(* IEC 61131-3 sources: kns-port-domestic/targets/astra/src/POUs/Model/F_PumpCurrent, 2 files *)

(* ---- F_PumpCurrent.decl.st ---- *)
// Назначение: ток двигателя насоса в модели, А. Гидравлическая мощность
//             P_hyd = ρ·g·(q/3600)·H/1000 кВт; потребляемая P = max(P_hyd/η, rLossShare·Pnom·s³) —
//             не меньше потерь без подачи, поэтому ток непрерывен при закрытии обратного клапана;
//             I = rImagShare·Inom·s + (1 − rImagShare)·Inom·P/Pnom. Без вращения (s ≤ 0), при
//             неверной характеристике или неконечных входах — 0.
// Автор:      kr0nsch
// Версия:     0.1.0
// Документ:   docs/DESIGN.md, разделы 11.2, 11.3
FUNCTION F_PumpCurrent : REAL
VAR_INPUT
    rFlow_m3h : REAL;           // подача насоса
    rHead_m   : REAL;           // напор сети в рабочей точке
    rSpeed    : REAL;           // относительная скорость s = f / 50 Гц
    stPump    : ST_PumpModelCfg;  // характеристика насоса и двигателя
END_VAR
VAR
    rHyd_kW  : REAL;            // гидравлическая мощность
    rLoss_kW : REAL;            // потери без подачи
    rIn_kW   : REAL;            // потребляемая мощность
END_VAR

(* ---- F_PumpCurrent.impl.st ---- *)
F_PumpCurrent := 0.0;
IF NOT (PL.F_IsFinite(rIn := rFlow_m3h) AND PL.F_IsFinite(rIn := rHead_m) AND PL.F_IsFinite(rIn := rSpeed)) THEN
    RETURN;
END_IF
IF rSpeed <= 0.0 OR stPump.rPnom_kW <= 0.0 OR stPump.rEta <= 0.0 THEN
    RETURN;
END_IF

rHyd_kW := GVL_Const.SIM_RHO_KGM3 * GVL_Const.SIM_GRAVITY_MPS2 * (MAX(rFlow_m3h, 0.0) / GVL_Const.SIM_S_PER_H)
           * MAX(rHead_m, 0.0) / GVL_Const.SIM_W_PER_KW;
rLoss_kW := stPump.rLossShare * stPump.rPnom_kW * rSpeed * rSpeed * rSpeed;
rIn_kW := MAX(rHyd_kW / stPump.rEta, rLoss_kW);
F_PumpCurrent := stPump.rImagShare * stPump.rInom_A * rSpeed
                 + (1.0 - stPump.rImagShare) * stPump.rInom_A * rIn_kW / stPump.rPnom_kW;
